//{attribute 'qualified_only'}
//{attribute 'strict'}
{attribute 'to_string'}
TYPE E_Recipe_Name :
(
	//e0_not_in_use := 0,
	R_All:=1,
	R_Device_Dough1,
	R_Device_Dough2,
	R_Device_Dough3,
	R_Device_Dough4,
	R_Piston_Settings // must be last
	
);
END_TYPE

(* stored: Version 1.1.0.1, ProductVersion 3.1.4024.12
   DUT E_Recipe_Name: Id {6073e4a2-137d-47fd-bf33-e5974ec005a2} *)
